(* IEC 61131-3 sources: llm-plc-st-eval/data/processed/gpt-4o/I5/few_shot, 3 files *)

(* ---- ejec_1.st ---- *)
FUNCTION_BLOCK FB_Clasificadora
VAR_INPUT
    sensorPresencia : BOOL; (* Sensor de presencia de piezas *)
    sensorAltura : BOOL;    (* Sensor de altura de piezas *)
END_VAR
VAR_OUTPUT
    banda : BOOL;           (* Banda transportadora activa *)
    piston : BOOL;          (* Pistón para desviar piezas altas *)
    nAltas : INT;           (* Contador de piezas altas *)
    nBajas : INT;           (* Contador de piezas bajas *)
END_VAR
VAR
    tRetraso : TON;         (* Temporizador de retraso de 2 segundos *)
    tPulso : TP;            (* Temporizador de pulso de 1 segundo *)
    piezaDetectada : BOOL;  (* Indica si una pieza ha sido detectada *)
END_VAR

(* La banda está siempre activa *)
banda := TRUE;

(* Detectar una pieza y verificar su altura *)
IF sensorPresencia AND NOT piezaDetectada THEN
    piezaDetectada := TRUE;
    IF sensorAltura THEN
        nAltas := nAltas + 1;
        tRetraso(IN := TRUE, PT := T#2S);
    ELSE
        nBajas := nBajas + 1;
    END_IF;
ELSIF NOT sensorPresencia THEN
    piezaDetectada := FALSE;
END_IF;

(* Activar el pistón después del retraso si la pieza es alta *)
IF tRetraso.Q THEN
    tPulso(IN := TRUE, PT := T#1S);
    tRetraso(IN := FALSE);
END_IF;

(* Salida del pistón controlada por el pulso de 1 segundo *)
piston := tPulso.Q;

END_FUNCTION_BLOCK

(* ---- ejec_2.st ---- *)
FUNCTION_BLOCK FB_Clasificadora
VAR_INPUT
    sensorPresencia : BOOL; (* Sensor de presencia de piezas *)
    sensorAltura : BOOL;    (* Sensor de altura de piezas *)
END_VAR
VAR_OUTPUT
    banda : BOOL;           (* Banda transportadora activa *)
    piston : BOOL;          (* Pistón para desviar piezas altas *)
    nAltas : INT;           (* Contador de piezas altas *)
    nBajas : INT;           (* Contador de piezas bajas *)
END_VAR
VAR
    tRetraso : TON;         (* Temporizador para retraso de 2 segundos *)
    tPulso : TON;           (* Temporizador para pulso de 1 segundo *)
    piezaAltaDetectada : BOOL; (* Indica si una pieza alta fue detectada *)
END_VAR

(* La banda transportadora siempre está activa *)
banda := TRUE;

(* Detectar pieza alta y activar temporizador de retraso *)
IF sensorPresencia AND sensorAltura THEN
    piezaAltaDetectada := TRUE;
    tRetraso(IN := TRUE, PT := T#2S);
ELSE
    tRetraso(IN := FALSE);
END_IF

(* Activar pistón después del retraso si una pieza alta fue detectada *)
IF tRetraso.Q THEN
    tPulso(IN := TRUE, PT := T#1S);
    IF NOT tPulso.Q THEN
        piston := TRUE;
    ELSE
        piston := FALSE;
        piezaAltaDetectada := FALSE; (* Resetear detección de pieza alta *)
        tPulso(IN := FALSE);
    END_IF
ELSE
    piston := FALSE;
END_IF

(* Contar piezas altas y bajas *)
IF sensorPresencia AND NOT sensorAltura THEN
    nBajas := nBajas + 1;
ELSIF sensorPresencia AND sensorAltura AND NOT piezaAltaDetectada THEN
    nAltas := nAltas + 1;
END_IF

END_FUNCTION_BLOCK

(* ---- ejec_3.st ---- *)
FUNCTION_BLOCK FB_Clasificadora
VAR_INPUT
    sensorPresencia : BOOL; (* Sensor de presencia de piezas *)
    sensorAltura : BOOL;    (* Sensor de altura de piezas *)
END_VAR
VAR_OUTPUT
    banda : BOOL;           (* Banda transportadora activa *)
    piston : BOOL;          (* Pistón para desviar piezas altas *)
    nAltas : INT;           (* Contador de piezas altas *)
    nBajas : INT;           (* Contador de piezas bajas *)
END_VAR
VAR
    tRetraso : TON;         (* Temporizador para retraso de 2 segundos *)
    tPulso : TON;           (* Temporizador para pulso de 1 segundo *)
    piezaAltaDetectada : BOOL; (* Indica si se detectó una pieza alta *)
END_VAR

(* La banda transportadora siempre está activa *)
banda := TRUE;

(* Detectar una pieza alta y activar el temporizador de retraso *)
IF sensorPresencia AND sensorAltura THEN
    piezaAltaDetectada := TRUE;
    tRetraso(IN := TRUE, PT := T#2S);
ELSE
    tRetraso(IN := FALSE);
END_IF

(* Activar el pistón 2 segundos después de detectar una pieza alta *)
IF tRetraso.Q THEN
    tPulso(IN := TRUE, PT := T#1S);
    piezaAltaDetectada := FALSE;
ELSE
    tPulso(IN := FALSE);
END_IF

(* Salida del pistón activa durante 1 segundo *)
piston := tPulso.Q;

(* Contar piezas altas y bajas *)
IF sensorPresencia AND NOT sensorAltura THEN
    nBajas := nBajas + 1;
ELSIF piezaAltaDetectada AND NOT tRetraso.Q THEN
    nAltas := nAltas + 1;
END_IF

END_FUNCTION_BLOCK
